Staubli VAL3: getLog.pgx

public program getLog(string& x_sLog[] (dimensions=1), num x_nType (dimensions=1))
begin
  call Log:getlog(x_sLog,x_nType)
end
